Fanuc KAREL source: kt00918.KL

PROGRAM KT00918
%NOLOCKGROUP
VAR
S1 : STRING[80];S2 : STRING[80];OUT:INTEGER
BEGIN
--
--
S1='A'
S2='B'
S1='A'
S2='B'
OUT=INDEX(S1,S1)
END KT00918
